KUKA KRL program: folge11.src, folge11.dat

--- folge11.src ---
&ACCESS RVP
&REL 1
&COMMENT bt2krl sim production Folge 11 plan 16#4F80
DEF FOLGE11()
   ; Generated by bt2krl 0.1.0 from bt2plc plan bt_1792076124_welding_cell_2_small (cell welding_cell_2_small), PLAN_ID 16#4F80
   ; Robot robot2 (R2), controller robot2, model KR240R2900_ULTRA, joint mapping identity
   ; Profile sim (bt2plc simulator telegram). NEVER install on a VW KS24 robot:
   ; its signals collide with the VW standard (Fertigmeldung, interlocks, PRG_NR).
   ; Do not edit: regenerate with bt2krl (plain KRL, no inline forms).
   ; Production Folge: 11 ops; per op: STEP, REQUEST, wait GRANT, delay, motion (exact stop at the end), hold, REQUEST := 0, wait GRANT released
   ;FOLD INI
      BAS(#INITMOV,0)
      $ADVANCE=3
      $APO.CPTP=100
   ;ENDFOLD
   ;FOLD PLAN ID 16#4F80
      IF BT_PLANL<>PLAN_ID THEN
         BT_ECODE=259
         BT_ERR=TRUE
         RETURN
      ENDIF
   ;ENDFOLD
   BT_RUN=TRUE
   ;FOLD START DEVIATION P1 1.0
      IF (ABS($AXIS_ACT.A1-P1.A1)>1.0) OR (ABS($AXIS_ACT.A2-P1.A2)>1.0) OR (ABS($AXIS_ACT.A3-P1.A3)>1.0) OR (ABS($AXIS_ACT.A4-P1.A4)>1.0) OR (ABS($AXIS_ACT.A5-P1.A5)>1.0) OR (ABS($AXIS_ACT.A6-P1.A6)>1.0) THEN
         BT_WCODE=513
      ENDIF
   ;ENDFOLD
   ;FOLD OP 1 W15 MASK 16#00000002
      ; zones IL02
      IF BT_ABRT THEN
         RETURN
      ENDIF
      BT_STEP=1
      $OUT[226]=TRUE ; REQ IL02
      WAIT FOR $IN[98] ; GRANT
      IF BT_ABRT THEN
         RETURN
      ENDIF
      BAS(#VEL_PTP,1)
      PTP P1 C_PTP
      BAS(#VEL_PTP,8)
      PTP P2 C_PTP
      BAS(#VEL_PTP,25)
      PTP P3 C_PTP
      BAS(#VEL_PTP,41)
      PTP P4 C_PTP
      BAS(#VEL_PTP,57)
      PTP P5 C_PTP
      BAS(#VEL_PTP,73)
      PTP P6 C_PTP
      BAS(#VEL_PTP,90)
      PTP P7 C_PTP
      BAS(#VEL_PTP,100)
      PTP P8 C_PTP
      PTP P9 C_PTP
      PTP P10 C_PTP
      BAS(#VEL_PTP,90)
      PTP P11 C_PTP
      BAS(#VEL_PTP,78)
      PTP P12 C_PTP
      BAS(#VEL_PTP,65)
      PTP P13 C_PTP
      BAS(#VEL_PTP,53)
      PTP P14 C_PTP
      BAS(#VEL_PTP,41)
      PTP P15 C_PTP
      BAS(#VEL_PTP,25)
      PTP P16 C_PTP
      BAS(#VEL_PTP,9)
      PTP P17 C_PTP
      BAS(#VEL_PTP,4)
      PTP P18 C_PTP
      BAS(#VEL_PTP,1)
      PTP P19
      WAIT SEC 0.5 ; hold
      $OUT[226]=FALSE ; RELEASE IL02
      WAIT FOR NOT $IN[98] ; GRANT released
   ;ENDFOLD
   ;FOLD OP 2 W14 MASK 16#00000001
      ; zones IL01
      IF BT_ABRT THEN
         RETURN
      ENDIF
      BT_STEP=2
      $OUT[225]=TRUE ; REQ IL01
      WAIT FOR $IN[97] ; GRANT
      IF BT_ABRT THEN
         RETURN
      ENDIF
      BAS(#VEL_PTP,4)
      PTP P20 C_PTP
      BAS(#VEL_PTP,8)
      PTP P21 C_PTP
      BAS(#VEL_PTP,23)
      PTP P22 C_PTP
      BAS(#VEL_PTP,38)
      PTP P23 C_PTP
      BAS(#VEL_PTP,52)
      PTP P24 C_PTP
      BAS(#VEL_PTP,61)
      PTP P25 C_PTP
      BAS(#VEL_PTP,45)
      PTP P26 C_PTP
      BAS(#VEL_PTP,30)
      PTP P27 C_PTP
      BAS(#VEL_PTP,15)
      PTP P28 C_PTP
      BAS(#VEL_PTP,5)
      PTP P29 C_PTP
      BAS(#VEL_PTP,1)
      PTP P30
      WAIT SEC 0.5 ; hold
      $OUT[225]=FALSE ; RELEASE IL01
      WAIT FOR NOT $IN[97] ; GRANT released
   ;ENDFOLD
   ;FOLD OP 3 W13 MASK 16#00000002
      ; zones IL02
      IF BT_ABRT THEN
         RETURN
      ENDIF
      BT_STEP=3
      $OUT[226]=TRUE ; REQ IL02
      WAIT FOR $IN[98] ; GRANT
      IF BT_ABRT THEN
         RETURN
      ENDIF
      BAS(#VEL_PTP,5)
      PTP P31 C_PTP
      BAS(#VEL_PTP,9)
      PTP P32 C_PTP
      BAS(#VEL_PTP,23)
      PTP P33 C_PTP
      BAS(#VEL_PTP,34)
      PTP P34 C_PTP
      BAS(#VEL_PTP,45)
      PTP P35 C_PTP
      BAS(#VEL_PTP,53)
      PTP P36 C_PTP
      BAS(#VEL_PTP,39)
      PTP P37 C_PTP
      BAS(#VEL_PTP,28)
      PTP P38 C_PTP
      BAS(#VEL_PTP,17)
      PTP P39 C_PTP
      BAS(#VEL_PTP,6)
      PTP P40 C_PTP
      BAS(#VEL_PTP,4)
      PTP P41 C_PTP
      BAS(#VEL_PTP,1)
      PTP P42
      WAIT SEC 0.5 ; hold
      $OUT[226]=FALSE ; RELEASE IL02
      WAIT FOR NOT $IN[98] ; GRANT released
   ;ENDFOLD
   ;FOLD OP 4 W10 MASK 16#00000001
      ; zones IL01
      IF BT_ABRT THEN
         RETURN
      ENDIF
      BT_STEP=4
      $OUT[225]=TRUE ; REQ IL01
      WAIT FOR $IN[97] ; GRANT
      IF BT_ABRT THEN
         RETURN
      ENDIF
      BAS(#VEL_PTP,4)
      PTP P43 C_PTP
      BAS(#VEL_PTP,1)
      PTP P44 C_PTP
      BAS(#VEL_PTP,13)
      PTP P45 C_PTP
      BAS(#VEL_PTP,27)
      PTP P46 C_PTP
      BAS(#VEL_PTP,13)
      PTP P47 C_PTP
      BAS(#VEL_PTP,4)
      PTP P48 C_PTP
      BAS(#VEL_PTP,1)
      PTP P49
      WAIT SEC 0.5 ; hold
      $OUT[225]=FALSE ; RELEASE IL01
      WAIT FOR NOT $IN[97] ; GRANT released
   ;ENDFOLD
   ;FOLD OP 5 W11 MASK 16#00000002
      ; zones IL02
      IF BT_ABRT THEN
         RETURN
      ENDIF
      BT_STEP=5
      $OUT[226]=TRUE ; REQ IL02
      WAIT FOR $IN[98] ; GRANT
      IF BT_ABRT THEN
         RETURN
      ENDIF
      BAS(#VEL_PTP,4)
      PTP P50 C_PTP
      BAS(#VEL_PTP,8)
      PTP P51 C_PTP
      BAS(#VEL_PTP,24)
      PTP P52 C_PTP
      BAS(#VEL_PTP,40)
      PTP P53 C_PTP
      BAS(#VEL_PTP,56)
      PTP P54 C_PTP
      BAS(#VEL_PTP,65)
      PTP P55 C_PTP
      BAS(#VEL_PTP,48)
      PTP P56 C_PTP
      BAS(#VEL_PTP,32)
      PTP P57 C_PTP
      BAS(#VEL_PTP,16)
      PTP P58 C_PTP
      BAS(#VEL_PTP,4)
      PTP P59 C_PTP
      BAS(#VEL_PTP,1)
      PTP P60
      WAIT SEC 0.5 ; hold
      $OUT[226]=FALSE ; RELEASE IL02
      WAIT FOR NOT $IN[98] ; GRANT released
   ;ENDFOLD
   ;FOLD OP 6 W12 MASK 16#00000001
      ; zones IL01
      IF BT_ABRT THEN
         RETURN
      ENDIF
      BT_STEP=6
      $OUT[225]=TRUE ; REQ IL01
      WAIT FOR $IN[97] ; GRANT
      IF BT_ABRT THEN
         RETURN
      ENDIF
      BAS(#VEL_PTP,5)
      PTP P61 C_PTP
      BAS(#VEL_PTP,9)
      PTP P62 C_PTP
      BAS(#VEL_PTP,25)
      PTP P63 C_PTP
      BAS(#VEL_PTP,42)
      PTP P64 C_PTP
      BAS(#VEL_PTP,55)
      PTP P65 C_PTP
      BAS(#VEL_PTP,65)
      PTP P66 C_PTP
      BAS(#VEL_PTP,50)
      PTP P67 C_PTP
      BAS(#VEL_PTP,34)
      PTP P68 C_PTP
      BAS(#VEL_PTP,17)
      PTP P69 C_PTP
      BAS(#VEL_PTP,4)
      PTP P70 C_PTP
      BAS(#VEL_PTP,1)
      PTP P71
      WAIT SEC 0.5 ; hold
      $OUT[225]=FALSE ; RELEASE IL01
      WAIT FOR NOT $IN[97] ; GRANT released
   ;ENDFOLD
   ;FOLD OP 7 ROBOT2_S06 MASK 16#00000002
      ; zones IL02
      IF BT_ABRT THEN
         RETURN
      ENDIF
      BT_STEP=7
      $OUT[226]=TRUE ; REQ IL02
      WAIT FOR $IN[98] ; GRANT
      IF BT_ABRT THEN
         RETURN
      ENDIF
      BAS(#VEL_PTP,4)
      PTP P72 C_PTP
      BAS(#VEL_PTP,8)
      PTP P73 C_PTP
      BAS(#VEL_PTP,24)
      PTP P74 C_PTP
      BAS(#VEL_PTP,40)
      PTP P75 C_PTP
      BAS(#VEL_PTP,51)
      PTP P76 C_PTP
      BAS(#VEL_PTP,63)
      PTP P77 C_PTP
      BAS(#VEL_PTP,75)
      PTP P78 C_PTP
      BAS(#VEL_PTP,83)
      PTP P79 C_PTP
      BAS(#VEL_PTP,94)
      PTP P80 C_PTP
      BAS(#VEL_PTP,100)
      PTP P81 C_PTP
      BAS(#VEL_PTP,98)
      PTP P82 C_PTP
      BAS(#VEL_PTP,87)
      PTP P83 C_PTP
      BAS(#VEL_PTP,75)
      PTP P84 C_PTP
      BAS(#VEL_PTP,67)
      PTP P85 C_PTP
      BAS(#VEL_PTP,55)
      PTP P86 C_PTP
      BAS(#VEL_PTP,44)
      PTP P87 C_PTP
      BAS(#VEL_PTP,32)
      PTP P88 C_PTP
      BAS(#VEL_PTP,20)
      PTP P89 C_PTP
      BAS(#VEL_PTP,8)
      PTP P90 C_PTP
      BAS(#VEL_PTP,1)
      PTP P91
      $OUT[226]=FALSE ; RELEASE IL02
      WAIT FOR NOT $IN[98] ; GRANT released
   ;ENDFOLD
   ;FOLD OP 8 ROBOT2_S07 MASK 16#00000001
      ; zones IL01
      IF BT_ABRT THEN
         RETURN
      ENDIF
      BT_STEP=8
      $OUT[225]=TRUE ; REQ IL01
      WAIT FOR $IN[97] ; GRANT
      IF BT_ABRT THEN
         RETURN
      ENDIF
      PTP P92
      WAIT SEC 0.05 ; step dwell
      $OUT[225]=FALSE ; RELEASE IL01
      WAIT FOR NOT $IN[97] ; GRANT released
   ;ENDFOLD
   ;FOLD OP 9 W09 MASK 16#00000002
      ; zones IL02
      IF BT_ABRT THEN
         RETURN
      ENDIF
      BT_STEP=9
      $OUT[226]=TRUE ; REQ IL02
      WAIT FOR $IN[98] ; GRANT
      IF BT_ABRT THEN
         RETURN
      ENDIF
      PTP P93 C_PTP
      BAS(#VEL_PTP,8)
      PTP P94 C_PTP
      BAS(#VEL_PTP,23)
      PTP P95 C_PTP
      BAS(#VEL_PTP,42)
      PTP P96 C_PTP
      BAS(#VEL_PTP,64)
      PTP P97 C_PTP
      BAS(#VEL_PTP,86)
      PTP P98 C_PTP
      BAS(#VEL_PTP,100)
      PTP P99 C_PTP
      BAS(#VEL_PTP,98)
      PTP P100 C_PTP
      BAS(#VEL_PTP,79)
      PTP P101 C_PTP
      BAS(#VEL_PTP,56)
      PTP P102 C_PTP
      BAS(#VEL_PTP,38)
      PTP P103 C_PTP
      BAS(#VEL_PTP,23)
      PTP P104 C_PTP
      BAS(#VEL_PTP,8)
      PTP P105 C_PTP
      BAS(#VEL_PTP,4)
      PTP P106 C_PTP
      BAS(#VEL_PTP,1)
      PTP P107
      WAIT SEC 0.5 ; hold
      $OUT[226]=FALSE ; RELEASE IL02
      WAIT FOR NOT $IN[98] ; GRANT released
   ;ENDFOLD
   ;FOLD OP 10 W07 MASK 16#00000001
      ; zones IL01
      IF BT_ABRT THEN
         RETURN
      ENDIF
      BT_STEP=10
      $OUT[225]=TRUE ; REQ IL01
      WAIT FOR $IN[97] ; GRANT
      IF BT_ABRT THEN
         RETURN
      ENDIF
      BAS(#VEL_PTP,4)
      PTP P108 C_PTP
      BAS(#VEL_PTP,9)
      PTP P109 C_PTP
      BAS(#VEL_PTP,23)
      PTP P110 C_PTP
      BAS(#VEL_PTP,36)
      PTP P111 C_PTP
      BAS(#VEL_PTP,49)
      PTP P112 C_PTP
      BAS(#VEL_PTP,62)
      PTP P113 C_PTP
      BAS(#VEL_PTP,80)
      PTP P114 C_PTP
      BAS(#VEL_PTP,98)
      PTP P115 C_PTP
      BAS(#VEL_PTP,85)
      PTP P116 C_PTP
      BAS(#VEL_PTP,71)
      PTP P117 C_PTP
      BAS(#VEL_PTP,58)
      PTP P118 C_PTP
      BAS(#VEL_PTP,45)
      PTP P119 C_PTP
      BAS(#VEL_PTP,27)
      PTP P120 C_PTP
      BAS(#VEL_PTP,9)
      PTP P121 C_PTP
      BAS(#VEL_PTP,4)
      PTP P122 C_PTP
      BAS(#VEL_PTP,1)
      PTP P123
      WAIT SEC 0.5 ; hold
      $OUT[225]=FALSE ; RELEASE IL01
      WAIT FOR NOT $IN[97] ; GRANT released
   ;ENDFOLD
   ;FOLD OP 11 HOME MASK 16#00000002
      ; zones IL02
      IF BT_ABRT THEN
         RETURN
      ENDIF
      BT_STEP=11
      $OUT[226]=TRUE ; REQ IL02
      WAIT FOR $IN[98] ; GRANT
      IF BT_ABRT THEN
         RETURN
      ENDIF
      BAS(#VEL_PTP,4)
      PTP P124 C_PTP
      BAS(#VEL_PTP,17)
      PTP P125 C_PTP
      BAS(#VEL_PTP,28)
      PTP P126 C_PTP
      BAS(#VEL_PTP,42)
      PTP P127 C_PTP
      BAS(#VEL_PTP,59)
      PTP P128 C_PTP
      BAS(#VEL_PTP,73)
      PTP P129 C_PTP
      BAS(#VEL_PTP,86)
      PTP P130 C_PTP
      BAS(#VEL_PTP,98)
      PTP P131 C_PTP
      BAS(#VEL_PTP,81)
      PTP P132 C_PTP
      BAS(#VEL_PTP,67)
      PTP P133 C_PTP
      BAS(#VEL_PTP,53)
      PTP P134 C_PTP
      BAS(#VEL_PTP,37)
      PTP P135 C_PTP
      BAS(#VEL_PTP,20)
      PTP P136 C_PTP
      BAS(#VEL_PTP,6)
      PTP P137
      $OUT[226]=FALSE ; RELEASE IL02
      WAIT FOR NOT $IN[98] ; GRANT released
   ;ENDFOLD
   ;FOLD FINISH
      WAIT SEC 0 ; advance-run stop
      BT_STEP=0
      BT_FIN=TRUE
      BT_RUN=FALSE
   ;ENDFOLD
END

--- folge11.dat ---
&ACCESS RVP
&REL 1
&COMMENT bt2krl sim data Folge 11 plan 16#4F80
DEFDAT FOLGE11
   ; Generated by bt2krl 0.1.0 from bt2plc plan bt_1792076124_welding_cell_2_small (cell welding_cell_2_small), PLAN_ID 16#4F80
   ; Robot robot2 (R2), controller robot2, model KR240R2900_ULTRA, joint mapping identity
   ; Profile sim (bt2plc simulator telegram). NEVER install on a VW KS24 robot:
   ; its signals collide with the VW standard (Fertigmeldung, interlocks, PRG_NR).
   ; Do not edit: regenerate with bt2krl (plain KRL, no inline forms).
   EXT BAS (BAS_COMMAND :IN,REAL :IN )
   DECL INT PLAN_ID=20352
   DECL AXIS P1={A1 0.0,A2 -90.0,A3 90.0,A4 0.0,A5 0.0,A6 0.0}
   DECL AXIS P2={A1 0.5737,A2 -89.9472,A3 89.956,A4 0.3877,A5 1.0443,A6 -1.071}
   DECL AXIS P3={A1 2.295,A2 -89.7886,A3 89.8242,A4 1.5508,A5 4.1772,A6 -4.2843}
   DECL AXIS P4={A1 5.1638,A2 -89.5242,A3 89.6045,A4 3.4894,A5 9.3988,A6 -9.6399}
   DECL AXIS P5={A1 9.1802,A2 -89.1541,A3 89.2968,A4 6.2035,A5 16.7092,A6 -17.1378}
   DECL AXIS P6={A1 14.3441,A2 -88.6783,A3 88.9013,A4 9.6931,A5 26.1082,A6 -26.7779}
   DECL AXIS P7={A1 20.6556,A2 -88.0967,A3 88.4179,A4 13.9581,A5 37.5959,A6 -38.5603}
   DECL AXIS P8={A1 24.2417,A2 -87.7663,A3 88.1433,A4 16.3813,A5 44.1231,A6 -45.255}
   DECL AXIS P9={A1 36.0758,A2 -86.6759,A3 87.2368,A4 24.3783,A5 65.6628,A6 -67.3472}
   DECL AXIS P10={A1 39.662,A2 -86.3455,A3 86.9622,A4 26.8016,A5 72.19,A6 -74.0419}
   DECL AXIS P11={A1 45.9736,A2 -85.7639,A3 86.4788,A4 31.0667,A5 83.6781,A6 -85.8246}
   DECL AXIS P12={A1 48.6991,A2 -85.5127,A3 86.27,A4 32.9085,A5 88.6388,A6 -90.9126}
   DECL AXIS P13={A1 53.2894,A2 -85.0898,A3 85.9184,A4 36.0103,A5 96.9937,A6 -99.4819}
   DECL AXIS P14={A1 55.1542,A2 -84.918,A3 85.7756,A4 37.2705,A5 100.3879,A6 -102.9632}
   DECL AXIS P15={A1 58.0231,A2 -84.6536,A3 85.5558,A4 39.2092,A5 105.6099,A6 -108.319}
   DECL AXIS P16={A1 59.7445,A2 -84.495,A3 85.424,A4 40.3724,A5 108.743,A6 -111.5326}
   DECL AXIS P17={A1 60.3184,A2 -84.4421,A3 85.3801,A4 40.7602,A5 109.7875,A6 -112.6039}
   DECL AXIS P18={A1 60.3184,A2 -84.0663,A3 89.4727,A4 39.8163,A5 106.378,A6 -115.6432}
   DECL AXIS P19={A1 60.3184,A2 -84.0663,A3 89.4727,A4 39.8163,A5 106.378,A6 -115.6432}
   DECL AXIS P20={A1 60.3185,A2 -84.4422,A3 85.38,A4 40.76,A5 109.7875,A6 -112.6038}
   DECL AXIS P21={A1 60.8906,A2 -84.5147,A3 85.1946,A4 39.7526,A5 109.5332,A6 -112.2067}
   DECL AXIS P22={A1 62.6056,A2 -84.7323,A3 84.6388,A4 36.7323,A5 108.7708,A6 -111.0161}
   DECL AXIS P23={A1 65.4635,A2 -85.0949,A3 83.7126,A4 31.6991,A5 107.5004,A6 -109.0321}
   DECL AXIS P24={A1 69.4644,A2 -85.6025,A3 82.416,A4 24.6532,A5 105.7219,A6 -106.2548}
   DECL AXIS P25={A1 76.4644,A2 -86.4906,A3 80.1475,A4 12.3255,A5 102.6103,A6 -101.3954}
   DECL AXIS P26={A1 79.8927,A2 -86.9255,A3 79.0364,A4 6.2879,A5 101.0863,A6 -99.0155}
   DECL AXIS P27={A1 82.178,A2 -87.2155,A3 78.2958,A4 2.2632,A5 100.0705,A6 -97.4291}
   DECL AXIS P28={A1 83.3203,A2 -87.3604,A3 77.9256,A4 0.2514,A5 99.5626,A6 -96.636}
   DECL AXIS P29={A1 83.463,A2 -87.7143,A3 82.7391,A4 0.0,A5 94.9753,A6 -96.5369}
   DECL AXIS P30={A1 83.463,A2 -87.7143,A3 82.7393,A4 0.0,A5 94.975,A6 -96.5369}
   DECL AXIS P31={A1 83.463,A2 -87.3785,A3 77.8794,A4 0.0,A5 99.4991,A6 -96.5369}
   DECL AXIS P32={A1 84.6918,A2 -87.2527,A3 78.4704,A4 -1.682,A5 99.5365,A6 -95.3447}
   DECL AXIS P33={A1 86.8764,A2 -87.0291,A3 79.5212,A4 -4.6727,A5 99.6029,A6 -93.225}
   DECL AXIS P34={A1 90.1535,A2 -86.6936,A3 81.0974,A4 -9.1588,A5 99.7026,A6 -90.0452}
   DECL AXIS P35={A1 94.5231,A2 -86.2462,A3 83.1992,A4 -15.1405,A5 99.8354,A6 -85.8055}
   DECL AXIS P36={A1 104.833,A2 -85.1909,A3 88.1583,A4 -29.2542,A5 100.1487,A6 -75.8019}
   DECL AXIS P37={A1 108.6568,A2 -84.7994,A3 89.9975,A4 -34.4887,A5 100.265,A6 -72.0917}
   DECL AXIS P38={A1 111.3882,A2 -84.5198,A3 91.3113,A4 -38.2277,A5 100.348,A6 -69.4415}
   DECL AXIS P39={A1 113.027,A2 -84.352,A3 92.0996,A4 -40.4713,A5 100.3978,A6 -67.8513}
   DECL AXIS P40={A1 113.5735,A2 -84.2961,A3 92.3624,A4 -41.2193,A5 100.4144,A6 -67.3211}
   DECL AXIS P41={A1 113.5735,A2 -83.434,A3 95.9948,A4 -40.7671,A5 97.0212,A6 -64.3387}
   DECL AXIS P42={A1 113.5735,A2 -83.4339,A3 95.9949,A4 -40.7671,A5 97.0212,A6 -64.3387}
   DECL AXIS P43={A1 113.5735,A2 -84.2961,A3 92.3625,A4 -41.2194,A5 100.4144,A6 -67.3211}
   DECL AXIS P44={A1 113.4743,A2 -84.2053,A3 92.2272,A4 -41.2464,A5 100.3807,A6 -67.425}
   DECL AXIS P45={A1 111.9902,A2 -82.8467,A3 90.2042,A4 -41.6508,A5 99.8755,A6 -68.9814}
   DECL AXIS P46={A1 106.7982,A2 -78.0936,A3 83.1267,A4 -43.0653,A5 98.1083,A6 -74.4261}
   DECL AXIS P47={A1 105.3153,A2 -76.736,A3 81.1052,A4 -43.4693,A5 97.6035,A6 -75.9811}
   DECL AXIS P48={A1 105.2165,A2 -76.0415,A3 84.7458,A4 -43.1814,A5 94.384,A6 -73.063}
   DECL AXIS P49={A1 105.2165,A2 -76.0415,A3 84.7458,A4 -43.1814,A5 94.384,A6 -73.063}
   DECL AXIS P50={A1 105.2164,A2 -76.6456,A3 80.9705,A4 -43.4959,A5 97.5699,A6 -76.0848}
   DECL AXIS P51={A1 104.6959,A2 -76.7137,A3 80.81,A4 -42.4209,A5 97.5045,A6 -76.5731}
   DECL AXIS P52={A1 103.1357,A2 -76.9179,A3 80.3289,A4 -39.1979,A5 97.3084,A6 -78.037}
   DECL AXIS P53={A1 100.5355,A2 -77.2581,A3 79.5272,A4 -33.8269,A5 96.9816,A6 -80.4765}
   DECL AXIS P54={A1 96.8954,A2 -77.7344,A3 78.4049,A4 -26.3079,A5 96.5241,A6 -83.8916}
   DECL AXIS P55={A1 90.5268,A2 -78.5679,A3 76.4412,A4 -13.1528,A5 95.7236,A6 -89.8667}
   DECL AXIS P56={A1 87.4077,A2 -78.976,A3 75.4794,A4 -6.71,A5 95.3316,A6 -92.793}
   DECL AXIS P57={A1 85.3285,A2 -79.2481,A3 74.8383,A4 -2.4151,A5 95.0703,A6 -94.7437}
   DECL AXIS P58={A1 84.2892,A2 -79.3841,A3 74.5179,A4 -0.2682,A5 94.9396,A6 -95.7188}
   DECL AXIS P59={A1 84.1594,A2 -79.4239,A3 78.9966,A4 0.0,A5 90.4272,A6 -95.8407}
   DECL AXIS P60={A1 84.1594,A2 -79.4239,A3 78.9966,A4 0.0,A5 90.4272,A6 -95.8407}
   DECL AXIS P61={A1 84.1594,A2 -79.4011,A3 74.478,A4 0.0,A5 94.9231,A6 -95.8407}
   DECL AXIS P62={A1 83.5658,A2 -79.127,A3 74.4456,A4 1.1295,A5 95.2311,A6 -96.3067}
   DECL AXIS P63={A1 81.7843,A2 -78.3044,A3 74.3488,A4 4.5193,A5 96.1549,A6 -97.7054}
   DECL AXIS P64={A1 78.8148,A2 -76.9332,A3 74.1875,A4 10.1698,A5 97.6947,A6 -100.0369}
   DECL AXIS P65={A1 76.8845,A2 -76.0419,A3 74.0828,A4 13.8428,A5 98.6956,A6 -101.5525}
   DECL AXIS P66={A1 69.9793,A2 -72.8534,A3 73.7078,A4 26.9822,A5 102.2762,A6 -106.974}
   DECL AXIS P67={A1 66.4146,A2 -71.2073,A3 73.5142,A4 33.7653,A5 104.1247,A6 -109.7729}
   DECL AXIS P68={A1 64.0379,A2 -70.1099,A3 73.3851,A4 38.2877,A5 105.3571,A6 -111.6389}
   DECL AXIS P69={A1 62.8493,A2 -69.561,A3 73.3205,A4 40.5495,A5 105.9735,A6 -112.5722}
   DECL AXIS P70={A1 62.7004,A2 -68.9133,A3 77.0333,A4 40.1152,A5 102.7791,A6 -115.5705}
   DECL AXIS P71={A1 62.7004,A2 -68.9132,A3 77.0335,A4 40.1152,A5 102.7789,A6 -115.5706}
   DECL AXIS P72={A1 62.7004,A2 -69.4922,A3 73.3127,A4 40.8329,A5 106.0505,A6 -112.6893}
   DECL AXIS P73={A1 62.1033,A2 -69.6875,A3 73.4714,A4 40.4441,A5 105.0409,A6 -111.6161}
   DECL AXIS P74={A1 60.3141,A2 -70.2728,A3 73.9476,A4 39.2789,A5 102.0146,A6 -108.4003}
   DECL AXIS P75={A1 57.3325,A2 -71.2479,A3 74.7411,A4 37.3371,A5 96.9715,A6 -103.0416}
   DECL AXIS P76={A1 55.3945,A2 -71.8818,A3 75.2569,A4 36.075,A5 93.6937,A6 -99.5586}
   DECL AXIS P77={A1 50.6243,A2 -73.442,A3 76.5265,A4 32.9685,A5 85.6254,A6 -90.9852}
   DECL AXIS P78={A1 47.7921,A2 -74.3684,A3 77.2803,A4 31.124,A5 80.835,A6 -85.895}
   DECL AXIS P79={A1 44.6553,A2 -75.3944,A3 78.1151,A4 29.0813,A5 75.5295,A6 -80.2573}
   DECL AXIS P80={A1 37.4994,A2 -77.7348,A3 80.0196,A4 24.4211,A5 63.4261,A6 -67.3963}
   DECL AXIS P81={A1 25.2007,A2 -81.7575,A3 83.2929,A4 16.4116,A5 42.6242,A6 -45.2923}
   DECL AXIS P82={A1 21.4737,A2 -82.9765,A3 84.2848,A4 13.9845,A5 36.3204,A6 -38.5939}
   DECL AXIS P83={A1 14.914,A2 -85.122,A3 86.0307,A4 9.7126,A5 25.2254,A6 -26.8045}
   DECL AXIS P84={A1 12.0759,A2 -86.0503,A3 86.786,A4 7.8643,A5 20.425,A6 -21.7035}
   DECL AXIS P85={A1 9.5418,A2 -86.8791,A3 87.4605,A4 6.214,A5 16.1388,A6 -17.1491}
   DECL AXIS P86={A1 5.3678,A2 -88.2443,A3 88.5714,A4 3.4957,A5 9.079,A6 -9.6473}
   DECL AXIS P87={A1 3.7279,A2 -88.7807,A3 89.0078,A4 2.4278,A5 6.3055,A6 -6.7001}
   DECL AXIS P88={A1 1.3425,A2 -89.5609,A3 89.6427,A4 0.8743,A5 2.2707,A6 -2.4128}
   DECL AXIS P89={A1 0.5969,A2 -89.8048,A3 89.8412,A4 0.3887,A5 1.0096,A6 -1.0727}
   DECL AXIS P90={A1 0.0001,A2 -90.0,A3 90.0,A4 0.0001,A5 0.0002,A6 -0.0002}
   DECL AXIS P91={A1 0.0,A2 -90.0,A3 90.0,A4 0.0,A5 0.0,A6 0.0}
   DECL AXIS P92={A1 0.0,A2 -90.0,A3 90.0,A4 0.0,A5 0.0,A6 0.0}
   DECL AXIS P93={A1 0.0,A2 -90.0,A3 90.0,A4 0.0,A5 0.0,A6 0.0}
   DECL AXIS P94={A1 0.5843,A2 -89.7203,A3 89.7053,A4 0.3797,A5 0.9612,A6 -0.9463}
   DECL AXIS P95={A1 2.337,A2 -88.8815,A3 88.821,A4 1.5187,A5 3.8445,A6 -3.785}
   DECL AXIS P96={A1 7.1569,A2 -86.5745,A3 86.3894,A4 4.6508,A5 11.7734,A6 -11.5913}
   DECL AXIS P97={A1 14.6063,A2 -83.0089,A3 82.6313,A4 9.4916,A5 24.0281,A6 -23.6565}
   DECL AXIS P98={A1 24.6855,A2 -78.1847,A3 77.5464,A4 16.0414,A5 40.6089,A6 -39.9809}
   DECL AXIS P99={A1 37.1096,A2 -72.2381,A3 71.2786,A4 24.1149,A5 61.047,A6 -60.103}
   DECL AXIS P100={A1 44.7047,A2 -68.6028,A3 67.4469,A4 29.0506,A5 73.5415,A6 -72.4043}
   DECL AXIS P101={A1 53.9067,A2 -64.1984,A3 62.8046,A4 35.0303,A5 88.6793,A6 -87.3079}
   DECL AXIS P102={A1 60.4798,A2 -61.0523,A3 59.4885,A4 39.3016,A5 99.4922,A6 -97.9536}
   DECL AXIS P103={A1 63.4012,A2 -59.654,A3 58.0147,A4 41.2001,A5 104.2981,A6 -102.6852}
   DECL AXIS P104={A1 65.1542,A2 -58.8149,A3 57.1304,A4 42.3392,A5 107.1818,A6 -105.5244}
   DECL AXIS P105={A1 65.7388,A2 -58.5351,A3 56.8355,A4 42.7191,A5 108.1435,A6 -106.4711}
   DECL AXIS P106={A1 65.7389,A2 -58.3151,A3 60.9792,A4 41.8475,A5 104.9144,A6 -109.5335}
   DECL AXIS P107={A1 65.7389,A2 -58.3151,A3 60.9793,A4 41.8474,A5 104.9142,A6 -109.5335}
   DECL AXIS P108={A1 65.7389,A2 -58.5351,A3 56.8356,A4 42.7191,A5 108.1435,A6 -106.4715}
   DECL AXIS P109={A1 66.2857,A2 -58.6182,A3 56.969,A4 41.5191,A5 108.0202,A6 -106.0735}
   DECL AXIS P110={A1 66.9695,A2 -58.7222,A3 57.136,A4 40.0185,A5 107.8658,A6 -105.576}
   DECL AXIS P111={A1 69.158,A2 -59.0548,A3 57.6706,A4 35.2157,A5 107.3716,A6 -103.9838}
   DECL AXIS P112={A1 70.6627,A2 -59.2834,A3 58.0382,A4 31.9136,A5 107.0318,A6 -102.8891}
   DECL AXIS P113={A1 74.4929,A2 -59.8656,A3 58.9739,A4 23.5079,A5 106.167,A6 -100.1025}
   DECL AXIS P114={A1 79.4176,A2 -60.614,A3 60.1769,A4 12.7002,A5 105.055,A6 -96.5196}
   DECL AXIS P115={A1 91.457,A2 -62.4437,A3 63.1179,A4 -13.7209,A5 102.3365,A6 -87.7606}
   DECL AXIS P116={A1 94.0567,A2 -62.8388,A3 63.753,A4 -19.4262,A5 101.7494,A6 -85.8692}
   DECL AXIS P117={A1 98.4353,A2 -63.5042,A3 64.8226,A4 -29.0353,A5 100.7607,A6 -82.6837}
   DECL AXIS P118={A1 100.2142,A2 -63.7746,A3 65.2571,A4 -32.9391,A5 100.3591,A6 -81.3895}
   DECL AXIS P119={A1 102.9509,A2 -64.1905,A3 65.9257,A4 -38.9453,A5 99.7411,A6 -79.3984}
   DECL AXIS P120={A1 104.5933,A2 -64.4402,A3 66.3269,A4 -42.5494,A5 99.3702,A6 -78.2035}
   DECL AXIS P121={A1 105.1411,A2 -64.5234,A3 66.4608,A4 -43.7516,A5 99.2465,A6 -77.805}
   DECL AXIS P122={A1 105.1412,A2 -64.0599,A3 70.284,A4 -43.3527,A5 96.139,A6 -74.8248}
   DECL AXIS P123={A1 105.1412,A2 -64.0599,A3 70.2842,A4 -43.3527,A5 96.1389,A6 -74.8246}
   DECL AXIS P124={A1 104.5586,A2 -64.2036,A3 70.3934,A4 -43.1125,A5 95.6061,A6 -74.41}
   DECL AXIS P125={A1 102.8102,A2 -64.635,A3 70.7213,A4 -42.3916,A5 94.0074,A6 -73.1657}
   DECL AXIS P126={A1 99.8957,A2 -65.354,A3 71.2678,A4 -41.1899,A5 91.3425,A6 -71.0916}
   DECL AXIS P127={A1 93.3377,A2 -66.972,A3 72.4976,A4 -38.4858,A5 85.346,A6 -66.4246}
   DECL AXIS P128={A1 84.1563,A2 -69.2373,A3 74.2192,A4 -34.7,A5 76.9506,A6 -59.8905}
   DECL AXIS P129={A1 76.5777,A2 -71.107,A3 75.6403,A4 -31.5752,A5 70.021,A6 -54.4972}
   DECL AXIS P130={A1 63.0236,A2 -74.451,A3 78.182,A4 -25.9864,A5 57.6275,A6 -44.8513}
   DECL AXIS P131={A1 37.3174,A2 -80.7932,A3 83.0023,A4 -15.387,A5 34.1222,A6 -26.5572}
   DECL AXIS P132={A1 24.636,A2 -83.9219,A3 85.3803,A4 -10.1581,A5 22.5267,A6 -17.5325}
   DECL AXIS P133={A1 17.6394,A2 -85.6481,A3 86.6923,A4 -7.2732,A5 16.129,A6 -12.5532}
   DECL AXIS P134={A1 9.3306,A2 -87.698,A3 88.2503,A4 -3.8473,A5 8.5317,A6 -6.6402}
   DECL AXIS P135={A1 3.6454,A2 -89.1006,A3 89.3164,A4 -1.5031,A5 3.3333,A6 -2.5943}
   DECL AXIS P136={A1 0.5837,A2 -89.856,A3 89.8905,A4 -0.2407,A5 0.5338,A6 -0.4154}
   DECL AXIS P137={A1 0.0,A2 -90.0,A3 90.0,A4 0.0,A5 0.0,A6 0.0}
ENDDAT
